// Characterization of FB_TelescopeControl (IAG50cm) for a stop during a slew, on mock axes (plan step 2, IAG50cmTests README).
// These tests pin what the code does today, with the line of the behaviour in a comment; they are not a specification. Every
// test owns a rig and runs over many PLC cycles (VAR_INST of the method, one Scan() per cycle); TcUnit calls all test methods
// every cycle, so the rigs warm up their clocks in parallel. A step that does not happen within its cycle budget fails the
// test with a message instead of hanging the run.
FUNCTION_BLOCK IagStopDuringSlew_Tests EXTENDS TcUnit.FB_TestSuite
VAR
END_VAR

Stop_During_Slew_One_Stop_For_The_Moving_Axis();
Stop_Drops_The_Move_Before_Sending_The_Axis_Stop();
Stop_Clears_The_Slew_And_Settles();

// #108: one MC_Stop per axis that is not at rest, none for an axis at rest. The IAG slew moves one axis at a time
// (_SlewTelescope stages 30..33 / 40..43), so only one axis is moving when the stop comes.
METHOD PRIVATE Stop_During_Slew_One_Stop_For_The_Moving_Axis
VAR_INST
	rig			: FB_IagRig;
	nStep		: INT;
	nCycles		: UINT;
	bHaMoving	: BOOL;
	sTest		: STRING(80);
END_VAR
TEST('Stop_During_Slew_One_Stop_For_The_Moving_Axis');
sTest := 'Stop_During_Slew_One_Stop_For_The_Moving_Axis: ';
IF nStep >= 90 THEN
	RETURN;
END_IF
rig.Scan();
nCycles := nCycles + 1;
CASE nStep OF
0:	// wait for the clock, then power on
	IF rig.ClockValid THEN
		rig.fbTel.Init();
		nStep := 10;
		nCycles := 0;
	ELSIF nCycles > 2000 THEN
		AssertTrue(Condition := FALSE, Message := 'the astronomical clock never became valid');
		F_Note(bFailed := NOT (FALSE), sText := CONCAT(sTest, 'the astronomical clock never became valid'));
		nStep := 99;
		TEST_FINISHED();
	END_IF
10:	// wait until the startup has finished (READY_STATE 1.0), then slew
	IF rig.Online THEN
		rig.fbTel.Slew(fAzimuth := 180.0, fAltitude := 45.0);
		nStep := 20;
		nCycles := 0;
	ELSIF nCycles > 1500 THEN
		AssertTrue(Condition := FALSE, Message := 'the mock telescope did not reach READY_STATE 1.0');
		F_Note(bFailed := NOT (FALSE), sText := CONCAT(sTest, 'the mock telescope did not reach READY_STATE 1.0'));
		nStep := 99;
		TEST_FINISHED();
	END_IF
20:	// wait until one axis is moving (the slew moves HA and Dec one after the other)
	IF rig.fbHa.MoveAxis OR rig.fbDec.MoveAxis THEN
		bHaMoving := rig.fbHa.MoveAxis;
		AssertTrue(Condition := rig.fbTel.bSlewActive, Message := 'bSlew is set while the slew runs');
		F_Note(bFailed := NOT (rig.fbTel.bSlewActive), sText := CONCAT(sTest, 'bSlew is set while the slew runs'));
		// IAG50cm#17 step 0.3: the coordinate chain runs inside the telescope (the migration must keep it running). The slew
		// target az 180 / alt 45 is on the meridian: Dec about latitude - 45 = 6.56 deg, hour angle about 0.
		AssertFalse(Condition := F_NoteNear(CONCAT(sTest, 'Julian date'), 2461000.0, rig.fbTel.fJd, 2000.0), Message := 'fJd follows the clock');
		AssertFalse(Condition := F_NoteNear(CONCAT(sTest, 'slew target Dec'), 51.5592378 - 45.0, rig.fbTel.fDeclinationCalc, 0.5), Message := 'slew target declination');
		AssertTrue(Condition := COS(rig.fbTel.fHourAngleCalc * 0.017453292519943295) > 0.9999, Message := 'slew target hour angle about 0');
		F_Note(bFailed := NOT (COS(rig.fbTel.fHourAngleCalc * 0.017453292519943295) > 0.9999), sText := CONCAT(sTest, 'slew target hour angle about 0'));
		AssertTrue(Condition := ABS(rig.fbTel.fDeclinationApparent) <= 90.0, Message := 'apparent declination is finite');
		F_Note(bFailed := NOT (ABS(rig.fbTel.fDeclinationApparent) <= 90.0), sText := CONCAT(sTest, 'apparent declination is finite'));
		AssertTrue(Condition := ABS(rig.fbTel.fElevationCalc) <= 90.0, Message := 'target elevation is finite');
		F_Note(bFailed := NOT (ABS(rig.fbTel.fElevationCalc) <= 90.0), sText := CONCAT(sTest, 'target elevation is finite'));
		nStep := 30;
		nCycles := 0;
	ELSIF nCycles > 300 THEN
		AssertTrue(Condition := FALSE, Message := 'the slew did not start an axis move');
		F_Note(bFailed := NOT (FALSE), sText := CONCAT(sTest, 'the slew did not start an axis move'));
		nStep := 99;
		TEST_FINISHED();
	END_IF
30:	// let the move run for a few scans, then stop
	IF nCycles >= 5 THEN
		rig.fbTel.Stop();
		nStep := 40;
		nCycles := 0;
	END_IF
40:	// wait until the stop has settled
	IF NOT rig.fbTel.bStopActive AND rig.fbTel.bStopped AND nCycles > 5 THEN
		AssertEquals_UINT(Expected := SEL(bHaMoving, UINT#0, UINT#1), Actual := rig.fbHa.nStopEdges, Message := 'HA: one stop if it was the moving axis, none otherwise');
		F_Note(bFailed := (SEL(bHaMoving, UINT#0, UINT#1)) <> (rig.fbHa.nStopEdges), sText := CONCAT(sTest, 'HA: one stop if it was the moving axis, none otherwise'));
		AssertEquals_UINT(Expected := SEL(bHaMoving, UINT#1, UINT#0), Actual := rig.fbDec.nStopEdges, Message := 'Dec: one stop if it was the moving axis, none otherwise');
		F_Note(bFailed := (SEL(bHaMoving, UINT#1, UINT#0)) <> (rig.fbDec.nStopEdges), sText := CONCAT(sTest, 'Dec: one stop if it was the moving axis, none otherwise'));
		nStep := 99;
		TEST_FINISHED();
	ELSIF nCycles > 400 THEN
		AssertTrue(Condition := FALSE, Message := 'the stop did not settle');
		F_Note(bFailed := NOT (FALSE), sText := CONCAT(sTest, 'the stop did not settle'));
		nStep := 99;
		TEST_FINISHED();
	END_IF
END_CASE
END_METHOD

// _StopTelescope (I:1927-1953): the first scan of a stop only drops MoveAxis (the first branch; that does not stop a running
// move); the axis stop (StopAxis) is sent in the next scan.
METHOD PRIVATE Stop_Drops_The_Move_Before_Sending_The_Axis_Stop
VAR_INST
	rig			: FB_IagRig;
	nStep		: INT;
	nCycles		: UINT;
	bHaMoving	: BOOL;
	sTest		: STRING(80);
END_VAR
TEST('Stop_Drops_The_Move_Before_Sending_The_Axis_Stop');
sTest := 'Stop_Drops_The_Move_Before_Sending_The_Axis_Stop: ';
IF nStep >= 90 THEN
	RETURN;
END_IF
rig.Scan();
nCycles := nCycles + 1;
CASE nStep OF
0:	// wait for the clock, then power on
	IF rig.ClockValid THEN
		rig.fbTel.Init();
		nStep := 10;
		nCycles := 0;
	ELSIF nCycles > 2000 THEN
		AssertTrue(Condition := FALSE, Message := 'the astronomical clock never became valid');
		F_Note(bFailed := NOT (FALSE), sText := CONCAT(sTest, 'the astronomical clock never became valid'));
		nStep := 99;
		TEST_FINISHED();
	END_IF
10:	// wait until the startup has finished (READY_STATE 1.0), then slew
	IF rig.Online THEN
		rig.fbTel.Slew(fAzimuth := 180.0, fAltitude := 45.0);
		nStep := 20;
		nCycles := 0;
	ELSIF nCycles > 1500 THEN
		AssertTrue(Condition := FALSE, Message := 'the mock telescope did not reach READY_STATE 1.0');
		F_Note(bFailed := NOT (FALSE), sText := CONCAT(sTest, 'the mock telescope did not reach READY_STATE 1.0'));
		nStep := 99;
		TEST_FINISHED();
	END_IF
20:	// wait until one axis is moving (the slew moves HA and Dec one after the other)
	IF rig.fbHa.MoveAxis OR rig.fbDec.MoveAxis THEN
		bHaMoving := rig.fbHa.MoveAxis;
		AssertTrue(Condition := rig.fbTel.bSlewActive, Message := 'bSlew is set while the slew runs');
		F_Note(bFailed := NOT (rig.fbTel.bSlewActive), sText := CONCAT(sTest, 'bSlew is set while the slew runs'));
		nStep := 30;
		nCycles := 0;
	ELSIF nCycles > 300 THEN
		AssertTrue(Condition := FALSE, Message := 'the slew did not start an axis move');
		F_Note(bFailed := NOT (FALSE), sText := CONCAT(sTest, 'the slew did not start an axis move'));
		nStep := 99;
		TEST_FINISHED();
	END_IF
30:	// let the move run for a few scans, then stop
	IF nCycles >= 5 THEN
		rig.fbTel.Stop();
		nStep := 40;
		nCycles := 0;
	END_IF
40:	// scan 1 of the stop has just run: the move is dropped, no axis stop yet; scan 2 sends it
	IF nCycles = 1 THEN
		AssertFalse(Condition := rig.fbHa.MoveAxis OR rig.fbDec.MoveAxis, Message := 'scan 1 of the stop drops the move');
		F_Note(bFailed := (rig.fbHa.MoveAxis OR rig.fbDec.MoveAxis), sText := CONCAT(sTest, 'scan 1 of the stop drops the move'));
		AssertFalse(Condition := rig.fbHa.StopAxis OR rig.fbDec.StopAxis, Message := 'scan 1 of the stop does not send an axis stop yet');
		F_Note(bFailed := (rig.fbHa.StopAxis OR rig.fbDec.StopAxis), sText := CONCAT(sTest, 'scan 1 of the stop does not send an axis stop yet'));
	ELSIF nCycles = 2 THEN
		AssertTrue(Condition := SEL(bHaMoving, rig.fbDec.StopAxis, rig.fbHa.StopAxis), Message := 'scan 2 sends the stop to the axis that was moving');
		F_Note(bFailed := NOT (SEL(bHaMoving, rig.fbDec.StopAxis, rig.fbHa.StopAxis)), sText := CONCAT(sTest, 'scan 2 sends the stop to the axis that was moving'));
		AssertFalse(Condition := SEL(bHaMoving, rig.fbHa.StopAxis, rig.fbDec.StopAxis), Message := 'scan 2 sends no stop to the axis at rest');
		F_Note(bFailed := (SEL(bHaMoving, rig.fbHa.StopAxis, rig.fbDec.StopAxis)), sText := CONCAT(sTest, 'scan 2 sends no stop to the axis at rest'));
		nStep := 99;
		TEST_FINISHED();
	END_IF
END_CASE
END_METHOD

// Arbitration (I:501-526): a user stop during a slew drops bSlew, runs the stop until the axes stand still, and releases bStop.
METHOD PRIVATE Stop_Clears_The_Slew_And_Settles
VAR_INST
	rig			: FB_IagRig;
	nStep		: INT;
	nCycles		: UINT;
	bHaMoving	: BOOL;
	sTest		: STRING(80);
END_VAR
TEST('Stop_Clears_The_Slew_And_Settles');
sTest := 'Stop_Clears_The_Slew_And_Settles: ';
IF nStep >= 90 THEN
	RETURN;
END_IF
rig.Scan();
nCycles := nCycles + 1;
CASE nStep OF
0:	// wait for the clock, then power on
	IF rig.ClockValid THEN
		rig.fbTel.Init();
		nStep := 10;
		nCycles := 0;
	ELSIF nCycles > 2000 THEN
		AssertTrue(Condition := FALSE, Message := 'the astronomical clock never became valid');
		F_Note(bFailed := NOT (FALSE), sText := CONCAT(sTest, 'the astronomical clock never became valid'));
		nStep := 99;
		TEST_FINISHED();
	END_IF
10:	// wait until the startup has finished (READY_STATE 1.0), then slew
	IF rig.Online THEN
		rig.fbTel.Slew(fAzimuth := 180.0, fAltitude := 45.0);
		nStep := 20;
		nCycles := 0;
	ELSIF nCycles > 1500 THEN
		AssertTrue(Condition := FALSE, Message := 'the mock telescope did not reach READY_STATE 1.0');
		F_Note(bFailed := NOT (FALSE), sText := CONCAT(sTest, 'the mock telescope did not reach READY_STATE 1.0'));
		nStep := 99;
		TEST_FINISHED();
	END_IF
20:	// wait until one axis is moving (the slew moves HA and Dec one after the other)
	IF rig.fbHa.MoveAxis OR rig.fbDec.MoveAxis THEN
		bHaMoving := rig.fbHa.MoveAxis;
		AssertTrue(Condition := rig.fbTel.bSlewActive, Message := 'bSlew is set while the slew runs');
		F_Note(bFailed := NOT (rig.fbTel.bSlewActive), sText := CONCAT(sTest, 'bSlew is set while the slew runs'));
		nStep := 30;
		nCycles := 0;
	ELSIF nCycles > 300 THEN
		AssertTrue(Condition := FALSE, Message := 'the slew did not start an axis move');
		F_Note(bFailed := NOT (FALSE), sText := CONCAT(sTest, 'the slew did not start an axis move'));
		nStep := 99;
		TEST_FINISHED();
	END_IF
30:	// let the move run for a few scans, then stop
	IF nCycles >= 5 THEN
		rig.fbTel.Stop();
		nStep := 40;
		nCycles := 0;
	END_IF
40:
	IF NOT rig.fbTel.bStopActive AND rig.fbTel.bStopped AND nCycles > 5 THEN
		AssertFalse(Condition := rig.fbTel.bSlewActive, Message := 'the stop dropped bSlew');
		F_Note(bFailed := (rig.fbTel.bSlewActive), sText := CONCAT(sTest, 'the stop dropped bSlew'));
		AssertFalse(Condition := rig.fbHa.MoveAxis OR rig.fbDec.MoveAxis, Message := 'no axis move is left');
		F_Note(bFailed := (rig.fbHa.MoveAxis OR rig.fbDec.MoveAxis), sText := CONCAT(sTest, 'no axis move is left'));
		AssertTrue(Condition := rig.fbTel.bReady, Message := 'the telescope is still ready after the stop');
		F_Note(bFailed := NOT (rig.fbTel.bReady), sText := CONCAT(sTest, 'the telescope is still ready after the stop'));
		nStep := 99;
		TEST_FINISHED();
	ELSIF nCycles > 400 THEN
		AssertTrue(Condition := FALSE, Message := 'the stop did not settle');
		F_Note(bFailed := NOT (FALSE), sText := CONCAT(sTest, 'the stop did not settle'));
		nStep := 99;
		TEST_FINISHED();
	END_IF
END_CASE
END_METHOD

END_FUNCTION_BLOCK

(* stored: Version 1.1.0.1, ProductVersion 3.1.4024.15
   POU IagStopDuringSlew_Tests: Id {5b3e06cb-4ef6-40a7-b073-cc1380feb139}, SpecialFunc None
   Method Stop_During_Slew_One_Stop_For_The_Moving_Axis: Id {aefa6ac1-f109-4163-a897-dbd0b91ae7dc}
   Method Stop_Drops_The_Move_Before_Sending_The_Axis_Stop: Id {c10fca0b-b98b-4f07-8436-58982a282ab0}
   Method Stop_Clears_The_Slew_And_Settles: Id {71f1a941-1613-44ee-bcb8-9d58e4de9677} *)
